(* PLC project SoftPN_Echo, Univision CODESYS CODESYS V3.5 SP22 Patch 4 *)
(* stored: creationDateTime 2026-10-19T14:30:00, modificationDateTime 2026-10-19T14:30:00 *)

PROGRAM PLC_PRG
  VAR
    abOut : ARRAY[0..31] OF BYTE;  (* PLC -> PC (Output 32 bytes): map in the module's I/O mapping, no AT *)
    abIn : ARRAY[0..31] OF BYTE;  (* PC -> PLC (Input 32 bytes): map in the module's I/O mapping, no AT *)
    tPattern : TON;
    bPattern : BYTE;  (* new pattern every 500 ms *)
    i : INT;
    dwHeartbeat : DWORD;  (* PC heartbeat, input bytes 0..3 (little-endian) *)
    dwLastBeat : DWORD;
    tSecond : TON;
    bHeartbeatOk : BOOL;  (* TRUE = the heartbeat changed during the last second: the PC is alive *)
    bEcho : BOOL;  (* TRUE = input bytes 4..31 equal output bytes 4..31 *)
    nEchoOk : UDINT;
    nEchoBad : UDINT;  (* small: one or two cycles of lag after each pattern change *)
  END_VAR

            // 1. write a pattern that changes every 500 ms into output bytes 4..31
tPattern(IN := NOT tPattern.Q, PT := T#500MS);
IF tPattern.Q THEN
    bPattern := bPattern + 1;
END_IF
FOR i := 4 TO 31 DO
    abOut[i] := bPattern + INT_TO_BYTE(i);
END_FOR

// 2. heartbeat counter written by the PC (input bytes 0..3, little-endian); must change every second
dwHeartbeat := SHL(BYTE_TO_DWORD(abIn[3]), 24) OR SHL(BYTE_TO_DWORD(abIn[2]), 16)
            OR SHL(BYTE_TO_DWORD(abIn[1]), 8) OR BYTE_TO_DWORD(abIn[0]);
tSecond(IN := NOT tSecond.Q, PT := T#1S);
IF tSecond.Q THEN
    bHeartbeatOk := dwHeartbeat <> dwLastBeat;
    dwLastBeat := dwHeartbeat;
END_IF

// 3. echo check: the PC copies our bytes 4..31 back
bEcho := TRUE;
FOR i := 4 TO 31 DO
    IF abIn[i] <> abOut[i] THEN
        bEcho := FALSE;
    END_IF
END_FOR
IF bEcho THEN
    nEchoOk := nEchoOk + 1;
ELSE
    nEchoBad := nEchoBad + 1;
END_IF
          
END_PROGRAM
